(* IEC 61131-3 sources: volt/packages/volt-lsp-iec/test-corpus/CodesysTestProject/Device/Plc Logic/Application/Library Manager/3SLicense, 22 files *)

(* ---- ACCESS_MODE.dut ---- *)
TYPE ACCESS_MODE :
(
	AM_READ,
	AM_WRITE,
	AM_APPEND,
	AM_READ_PLUS,
	AM_WRITE_PLUS,
	AM_APPEND_PLUS
);
END_TYPE

(* ---- CMPMGR_LICENSEREQUEST.dut ---- *)
TYPE CMPMGR_LICENSEREQUEST :
STRUCT
	ULLICENSEID : UDINT;
	ULLICENSEVALUE : UDINT;
END_STRUCT
END_TYPE

(* ---- RTS_CMBOXENTRY.dut ---- *)
TYPE RTS_CMBOXENTRY :
STRUCT
	MUSBOXMASK : WORD;
	MULBOXSERIAL : UDINT;
	MFLFICTRL : UDINT;
	MULFIRMCODE : UDINT;
	MUSFIRMACCESSCOUNTER : WORD;
	MUSFIRMITEMREF : WORD;
	MULFIRMUPDATECOUNTER : UDINT;
	MULFIRMPRECISETIME : UDINT;
	MAUSFIRMITEMTEXT : WSTRING(255);
	MULPRODUCTCODE : UDINT;
	MULFEATUREMAP : UDINT;
	MULUNITCOUNTER : UDINT;
	MULLICENSEQUANTITY : UDINT;
	MUSPRODUCTITEMREF : WORD;
END_STRUCT
END_TYPE

(* ---- EVENTIDS.gvl ---- *)
VAR_GLOBAL
	CMPMGR_LICENSEREQUEST : WORD := 16#1;
END_VAR

(* ---- GVL_HIDDEN.gvl ---- *)
VAR_GLOBAL
	GC_UIMAXFILESIZE : UINT := 512;
	GC_UIMAXSTOREDLIC : UINT := 64;
	GC_CLASSID_LICENSE : UDINT := 16#100D;
	GC_TDEMO : TIME := TIME#120m0s0ms;
	GC_TCYCLE : TIME := TIME#1m0s0ms;
	GC_TRESYNC : TIME := TIME#2s0ms;
	G_TDEMOTIME : TIME := TIME#120m0s0ms;
	G_OLM : OLM_OnlineLicenseManager;
	G_UDISTART : DWORD;
END_VAR

(* ---- CODEMGETCONTENTBYFIRMCODE_LOCAL.pou ---- *)
FUNCTION CODEMGETCONTENTBYFIRMCODE_LOCAL : RTS_IEC_RESULT
VAR_INPUT
	DUIFIRMCODE : UDINT;
	DUIPRODUCTCODE : UDINT;
END_VAR
VAR_IN_OUT
	LICENSEENTRY : RTS_CMBOXENTRY;
END_VAR
END_FUNCTION

(* ---- CODEMGETFEATUREMAPBYFIRMCODE_LOCAL.pou ---- *)
FUNCTION CODEMGETFEATUREMAPBYFIRMCODE_LOCAL : UDINT
VAR_INPUT
	DUIFIRMCODE : UDINT;
	DUIPRODUCTCODE : UDINT;
END_VAR
END_FUNCTION

(* ---- FCTCONFDYNLICCHALLENGE.pou ---- *)
FUNCTION FCTCONFDYNLICCHALLENGE : BOOL
VAR_INPUT
	UDILICENSEID : UDINT;
	UDINEWLICENSEVALUE : UDINT;
	UDICHALLENGE : UDINT;
	PRESULT : POINTER TO RTS_IEC_RESULT;
END_VAR
END_FUNCTION

(* ---- FCTGETUSERLICENSEVALUE.pou ---- *)
FUNCTION FCTGETUSERLICENSEVALUE : UDINT
VAR_INPUT
	UDILICENSEID : UDINT;
	PRESULT : POINTER TO RTS_IEC_RESULT;
END_VAR
END_FUNCTION

(* ---- FCTREQDYNLICCHALLENGE.pou ---- *)
FUNCTION FCTREQDYNLICCHALLENGE : UDINT
VAR_INPUT
	UDILICENSEID : UDINT;
	UDINEWLICENSEVALUE : UDINT;
	PRESULT : POINTER TO RTS_IEC_RESULT;
END_VAR
END_FUNCTION

(* ---- MYSTRING_TO_UDINT.pou ---- *)
FUNCTION MYSTRING_TO_UDINT : UDINT
VAR_INPUT
	STR : STRING;
END_VAR
END_FUNCTION

(* ---- MYUDINT_TO_STRING.pou ---- *)
FUNCTION MYUDINT_TO_STRING : STRING(10)
VAR_INPUT
	UDI : UDINT;
END_VAR
END_FUNCTION

(* ---- REGISTERLICENSEFUNCTIONS.pou ---- *)
FUNCTION REGISTERLICENSEFUNCTIONS : RTS_IEC_RESULT
END_FUNCTION

(* ---- SYSFILECLOSE.pou ---- *)
FUNCTION SYSFILECLOSE : RTS_IEC_RESULT
VAR_INPUT
	HFILE : RTS_IEC_HANDLE;
END_VAR
END_FUNCTION

(* ---- SYSFILEGETSIZEBYHANDLE.pou ---- *)
FUNCTION SYSFILEGETSIZEBYHANDLE : __XWORD
VAR_INPUT
	HFILE : RTS_IEC_HANDLE;
	PRESULT : POINTER TO RTS_IEC_RESULT;
END_VAR
END_FUNCTION

(* ---- SYSFILEOPEN.pou ---- *)
FUNCTION SYSFILEOPEN : RTS_IEC_HANDLE
VAR_INPUT
	SZFILE : REFERENCE TO STRING;
	AM : ACCESS_MODE;
	PRESULT : POINTER TO RTS_IEC_RESULT;
END_VAR
END_FUNCTION

(* ---- SYSFILEREAD.pou ---- *)
FUNCTION SYSFILEREAD : __XWORD
VAR_INPUT
	HFILE : RTS_IEC_HANDLE;
	PBYBUFFER : POINTER TO BYTE;
	ULSIZE : __XWORD;
	PRESULT : POINTER TO RTS_IEC_RESULT;
END_VAR
END_FUNCTION

(* ---- SYSTARGETGETID.pou ---- *)
FUNCTION SYSTARGETGETID : RTS_IEC_RESULT
VAR_INPUT
	PULTARGETID : POINTER TO DWORD;
END_VAR
END_FUNCTION

(* ---- SYSTARGETGETTYPE.pou ---- *)
FUNCTION SYSTARGETGETTYPE : RTS_IEC_RESULT
VAR_INPUT
	PULTYPE : POINTER TO DWORD;
END_VAR
END_FUNCTION

(* ---- UNREGISTERLICENSEFUNCTIONS.pou ---- *)
FUNCTION UNREGISTERLICENSEFUNCTIONS : RTS_IEC_RESULT
END_FUNCTION

(* ---- OLM_COMMCYCLE.pou ---- *)
FUNCTION_BLOCK OLM_COMMCYCLE
VAR
	_TLASTCYCLE : TIME := TIME();
END_VAR
END_FUNCTION_BLOCK

METHOD EVENTCALLBACK : SysTypes.RTS_IEC_RESULT
VAR_INPUT
	PEVENTPARAM : POINTER TO EventParam;
END_VAR
END_METHOD

(* ---- OLM_ONLINELICENSEMANAGER.pou ---- *)
FUNCTION_BLOCK OLM_ONLINELICENSEMANAGER
VAR
	_HFILE : RTS_IEC_HANDLE;
	_UDITARGET : UDINT;
	_UDITYPE : UDINT;
	_UDICPU : UDINT;
	_UDIOS : UDINT;
	_ABYFILECONTENT : ARRAY [1..gc_uiMaxFileSize] OF BYTE;
	_UIFILESIZE : UINT;
	_XFILEREAD : BOOL;
	_UISTOREDLICENSES : UINT;
	_UDIDYNLICREQID : UDINT;
	_UDIDYNLICREQVALUE : UDINT;
	_UDIDYNLICCHALLENGE : UDINT;
	_XDEMOMESSAGE : BOOL;
	_SEMASTORE : UDINT;
	_LWLICENSEEVENTSENT : ULINT;
	_ADWLICENSESSTORED : ARRAY [1..gc_uiMaxStoredLic] OF ARRAY [1..3] OF DWORD;
	_HCYCLEEVENT : RTS_IEC_HANDLE;
	_HCYCLECALLBACK : RTS_IEC_HANDLE;
	_CCFB : OLM_CommCycle;
	_UIRESYNCSTOREDLICENSES : UINT;
	_UILASTRESYNCSTOREDLICENSES : UINT;
	_DWRESYNCLICNEXT : DWORD;
	_XRESYNCINIT : BOOL;
	_XRESYNCRECALL : BOOL;
END_VAR
END_FUNCTION_BLOCK

METHOD CODEMGETCONTENTBYFIRMCODE : RTS_IEC_RESULT
VAR_INPUT
	DUIFIRMCODE : UDINT;
	DUIPRODUCTCODE : UDINT;
END_VAR
VAR_IN_OUT
	LICENSEENTRY : RTS_CMBOXENTRY;
END_VAR
END_METHOD

METHOD CONFDYNLICCHALLENGE : BOOL
VAR_INPUT
	UDILICENSEID : UDINT;
	UDINEWLICENSEVALUE : UDINT;
	UDICHALLENGE : UDINT;
END_VAR
END_METHOD

METHOD CYCLICRESYNCCHECK
END_METHOD

METHOD DEMOMODEEXPIRED
VAR_INPUT
	STRCOMPONENT : STRING;
END_VAR
END_METHOD

METHOD DEMOMODEEXPIREDID
VAR_INPUT
	STRCOMPONENT : STRING;
	UDILICENSEID : UDINT;
END_VAR
END_METHOD

METHOD DEMOMODESTARTED
VAR_INPUT
	STRCOMPONENT : STRING;
END_VAR
END_METHOD

METHOD DEMOMODESTARTEDID
VAR_INPUT
	STRCOMPONENT : STRING;
	UDILICENSEID : UDINT;
END_VAR
END_METHOD

METHOD GENERATEEXCEPTION
END_METHOD

METHOD GETCODEMETERLICENSEVALUE : UDINT
VAR_INPUT
	UDIPRODUCTCODE : UDINT;
END_VAR
END_METHOD

METHOD GETDEMOLICENSE : UDINT
END_METHOD

METHOD GETLICENSEVALUE : UDINT
VAR_INPUT
	UDILICENSEID : UDINT;
END_VAR
END_METHOD

METHOD GETLICENSEVALUEBIT : INT
VAR_INPUT
	UDILICENSEID : UDINT;
	USIBIT : USINT;
END_VAR
END_METHOD

METHOD GETPURELICENSEVALUE : UDINT
VAR_INPUT
	UDILICENSEID : UDINT;
	XNOTFROMCACHE : BOOL;
END_VAR
VAR_OUTPUT
	UIPOSINCACHE : UINT;
END_VAR
END_METHOD

METHOD GETUSERLICENSEVALUE : UDINT
VAR_INPUT
	UDILICENSEID : UDINT;
END_VAR
END_METHOD

METHOD LICENSEMISSING
VAR_INPUT
	STRCOMPONENT : STRING;
END_VAR
END_METHOD

METHOD LICENSEMISSINGID
VAR_INPUT
	STRCOMPONENT : STRING;
	UDILICENSEID : UDINT;
END_VAR
END_METHOD

METHOD LOGERRORMESSAGE
VAR_INPUT
	STR : STRING;
END_VAR
END_METHOD

METHOD LOGINFOMESSAGE
VAR_INPUT
	STR : STRING;
END_VAR
END_METHOD

METHOD READLICENSEFILE : BOOL
END_METHOD

METHOD REQDYNLICCHALLENGE : UDINT
VAR_INPUT
	UDILICENSEID : UDINT;
	UDINEWLICENSEVALUE : UDINT;
END_VAR
END_METHOD

METHOD RESYNCLICENSEVALUES : BOOL
END_METHOD

METHOD STORELICENSE : UINT
VAR_INPUT
	UDILICENSEID : UDINT;
	UDIVALUE : UDINT;
END_VAR
END_METHOD

METHOD UDINTVALUEOFLINE : UDINT
VAR_INPUT
	STRID : STRING;
END_VAR
END_METHOD

METHOD VALUEOFLINE : STRING
VAR_INPUT
	STRID : STRING;
END_VAR
END_METHOD

METHOD FB_EXIT : BOOL
VAR_INPUT
	BINCOPYCODE : BOOL;
END_VAR
END_METHOD

METHOD FB_INIT : BOOL
VAR_INPUT
	BINITRETAINS : BOOL;
	BINCOPYCODE : BOOL;
END_VAR
END_METHOD

METHOD SENDEVENT
VAR_INPUT
	ULLICENSEID : UDINT;
	ULLICENSEVALUE : UDINT;
END_VAR
END_METHOD
